(* IEC 61131-3 sources: plc-st-test/packages/ingestors/generic/test/fixtures/plain/src, 1 file *)

(* ---- FB_A.st ---- *)
FUNCTION_BLOCK FB_A
VAR
  x : INT;
END_VAR
x := 1;
END_FUNCTION_BLOCK
